// TIA Portal V20 export
Screen "150PRBCompleteDisplay_3"  1276x673
  ScreenItem "Title_ScreenOverview_X390_Y2" at 390,2 size 500x30  Type=HmiTextBox
  ScreenItem "Button_Back_1" at 2,2 size 90x60  Type=HmiButton
  ScreenItem "sequenceControlFaceplate_Lite_1" at 357,556 size 641x64  Type=HmiFaceplateContainer
  ScreenItem "Line_Header_X0_Y64" at 82,780 size 1276x0  Type=HmiLine
  ScreenItem "permanentareaborderrectangle" at 0,0 size 0x0  Type=HmiRectangle
  ScreenItem "Button_Back" at 2,4 size 90x60  Type=HmiButton
  ScreenItem "Title_ScreenOverview_X390_Y2_1" at 380,5 size 510x57  Type=HmiTextBox
  ScreenItem "Line_Header_X0_Y64_1" at 0,64 size 1276x0  Type=HmiLine
  ScreenItem "面板容器_6" at 699,264 size 163x70  Type=HmiFaceplateContainer
  ScreenItem "面板容器_5" at 883,264 size 163x70  Type=HmiFaceplateContainer
  ScreenItem "面板容器_7" at 699,332 size 163x70  Type=HmiFaceplateContainer
  ScreenItem "面板容器_3" at 285,267 size 163x70  Type=HmiFaceplateContainer
  ScreenItem "面板容器_1" at 102,267 size 163x70  Type=HmiFaceplateContainer
  ScreenItem "面板容器_4" at 102,335 size 163x70  Type=HmiFaceplateContainer
  ScreenItem "Move_Legend" at 1182,2 size 90x60  Type=HmiButton
  ScreenItem "面板容器_2" at 1090,4 size 88x58  Type=HmiFaceplateContainer
  ScreenItem "OPMode1_Blocked" at 1164,6 size 14x14  Type=HmiGraphicView
  ScreenItem "OPMode4_Foreground_Blocked" at 1090,4 size 88x58  Type=HmiGraphicView
